// TIA Portal V20 export
// export: Created 2026-11-12T08:00:00.0000000Z, ExportSetting None, DisplayName Totally Integrated Automation Portal, DisplayVersion V20, DisplayName STEP 7 Professional, DisplayVersion V20
FUNCTION_BLOCK "FB_Valve_TonDelay_Pulse_LAD"   // FB22, LAD
TITLE = FB_Valve_TonDelay_Pulse_LAD
{ S7_Optimized_Access := 'TRUE' }
// 电磁阀单周期触发脉冲与通电延时确认（TON_TIME + PBox Static 边沿保持）
// stored: AutoNumber false, MemoryReserve 50, SetENOAutomatically false
   VAR_INPUT
      enable : Bool;
      triggerCmd : Bool;
      eStopNC : Bool;
      presetDelay : Time;
   END_VAR
   VAR_OUTPUT
      valveOut : Bool;
      triggerPulse : Bool;
      delayDone : Bool;
   END_VAR
   VAR
      statPrevEdge : Bool;
      tonInst { S7_SetPoint := 'True'} : TON_TIME;
   END_VAR
   VAR_TEMP   // added for the SCL form of the ladder/FBD networks
      _w1 : Bool;
      _w2 : Bool;
   END_VAR
BEGIN

REGION Network 1: 触发单脉冲检测
   // 网络1：在使能与急停正常后检测触发指令上升沿，输出单扫描周期脉冲
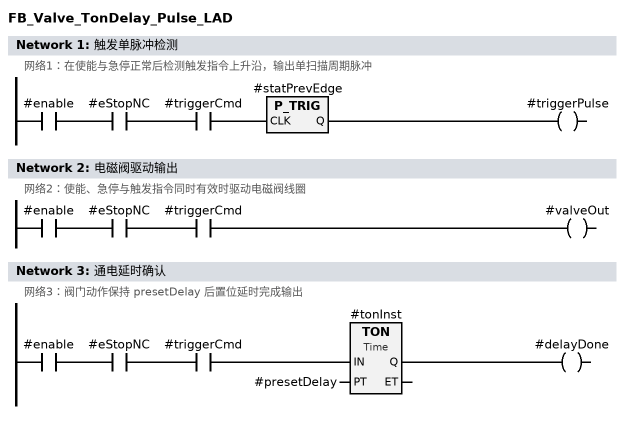
   RUNG wire#powerrail
      Contact( #enable )
      Contact( #eStopNC )
      Contact( #triggerCmd )
      P_Trig( #statPrevEdge )
      Coil( #triggerPulse )
   END_RUNG
   // the same network as SCL:
   #_w1 := #enable AND #eStopNC AND #triggerCmd;
   #_w2 := #_w1 AND NOT #statPrevEdge;   // rising edge
   #statPrevEdge := #_w1;
   #triggerPulse := #_w2;
END_REGION

REGION Network 2: 电磁阀驱动输出
   // 网络2：使能、急停与触发指令同时有效时驱动电磁阀线圈
   RUNG wire#powerrail
      Contact( #enable )
      Contact( #eStopNC )
      Contact( #triggerCmd )
      Coil( #valveOut )
   END_RUNG
   // the same network as SCL:
   #valveOut := #enable AND #eStopNC AND #triggerCmd;
END_REGION

REGION Network 3: 通电延时确认
   // 网络3：阀门动作保持 presetDelay 后置位延时完成输出
   RUNG wire#powerrail
      Contact( #enable )
      Contact( #eStopNC )
      Contact( #triggerCmd )
      { S7_Templates := "time_type := Time" } #tonInst.TON(pt := #presetDelay, et =>)
      Coil( #delayDone )
   END_RUNG
   // the same network as SCL:
   #tonInst(IN := #enable AND #eStopNC AND #triggerCmd, PT := #presetDelay);   // TON
   #delayDone := #tonInst.Q;
END_REGION
END_FUNCTION_BLOCK
